// TIA Portal V20 export
// export: Created 2026-10-12T16:46:22.2661913Z, ExportSetting WithDefaults, DisplayName Totally Integrated Automation Portal, DisplayVersion V20 Update 6, DisplayName TIA Portal Openness, DisplayVersion V20 Update 6, DisplayName TIA Portal Version Control Interface, DisplayVersion V20 Update 6, DisplayName SINAMICS Startdrive Advanced, DisplayVersion V20 SP1 Update 2, DisplayName SINAMICS Startdrive G110M, G120, G120C, G120D, G120P, G115D, DisplayVersion V20 SP1 Update 2, DisplayName SINAMICS Startdrive G130, G150, S120, S150, SINAMICS MV, G220, S200, S210, DisplayVersion V20 SP1 Update 2, DisplayName STEP 7 Professional, DisplayVersion V20 Update 6, DisplayName STEP 7 Safety, DisplayVersion V20 Update 2, DisplayName WinCC Basic/Comfort/Advanced, DisplayVersion V20 Update 6, DisplayName WinCC Professional, DisplayVersion V20 Update 6, DisplayName WinCC Unified, DisplayVersion V20 Update 6
VAR_GLOBAL   // PLC tag table "KP8"
   "Maschinenleuchte orange ein P01" AT %Q1001.4 : Bool;
   "Maschinenleuchte gruen ein P01" AT %Q1001.5 : Bool;
   "Maschinenleuchte rot ein P01" AT %Q1001.6 : Bool;
   "Maschinenleuchte orange ein P02" AT %Q2001.4 : Bool;
   "Maschinenleuchte gruen ein P02" AT %Q2001.5 : Bool;
   "Maschinenleuchte rot ein P02" AT %Q2001.6 : Bool;
   "Maschinenleuchte orange ein P03" AT %Q3001.4 : Bool;
   "Maschinenleuchte gruen ein P03" AT %Q3001.5 : Bool;
   "Maschinenleuchte rot ein P03" AT %Q3001.6 : Bool;
   "Maschinenleuchte orange ein P04" AT %Q4001.4 : Bool;
   "Maschinenleuchte gruen ein P04" AT %Q4001.5 : Bool;
   "Maschinenleuchte rot ein P04" AT %Q4001.6 : Bool;
   "Maschinenleuchte orange ein P05" AT %Q5001.4 : Bool;
   "Maschinenleuchte gruen ein P05" AT %Q5001.5 : Bool;
   "Maschinenleuchte rot ein P05" AT %Q5001.6 : Bool;
   "Maschinenleuchte orange ein P06" AT %Q6001.4 : Bool;
   "Maschinenleuchte gruen ein P06" AT %Q6001.5 : Bool;
   "Maschinenleuchte rot ein P06" AT %Q6001.6 : Bool;
   "Maschinenleuchte orange ein P07" AT %Q7001.4 : Bool;
   "Maschinenleuchte gruen ein P07" AT %Q7001.5 : Bool;
   "Maschinenleuchte rot ein P07" AT %Q7001.6 : Bool;
   "Maschinenleuchte orange ein P08" AT %Q8001.4 : Bool;
   "Maschinenleuchte gruen ein P08" AT %Q8001.5 : Bool;
   "Maschinenleuchte rot ein P08" AT %Q8001.6 : Bool;
   "Maschinenleuchte orange ein P09" AT %Q9001.4 : Bool;
   "Maschinenleuchte gruen ein P09" AT %Q9001.5 : Bool;
   "Maschinenleuchte rot ein P09" AT %Q9001.6 : Bool;
   "Maschinenleuchte orange ein P10" AT %Q10001.4 : Bool;
   "Maschinenleuchte gruen ein P10" AT %Q10001.5 : Bool;
   "Maschinenleuchte rot ein P10" AT %Q10001.6 : Bool;
   "Maschinenleuchte orange ein P11" AT %Q11001.4 : Bool;
   "Maschinenleuchte gruen ein P11" AT %Q11001.5 : Bool;
   "Maschinenleuchte rot ein P11" AT %Q11001.6 : Bool;
   "Maschinenleuchte orange ein P12" AT %Q12001.4 : Bool;
   "Maschinenleuchte gruen ein P12" AT %Q12001.5 : Bool;
   "Maschinenleuchte rot ein P12" AT %Q12001.6 : Bool;
   "Maschinenleuchte orange ein P13" AT %Q13001.4 : Bool;
   "Maschinenleuchte gruen ein P13" AT %Q13001.5 : Bool;
   "Maschinenleuchte rot ein P13" AT %Q13001.6 : Bool;
   "Maschinenleuchte orange ein P14" AT %Q14001.4 : Bool;
   "Maschinenleuchte gruen ein P14" AT %Q14001.5 : Bool;
   "Maschinenleuchte rot ein P14" AT %Q14001.6 : Bool;
   "Maschinenleuchte orange ein P15" AT %Q15001.4 : Bool;
   "Maschinenleuchte gruen ein P15" AT %Q15001.5 : Bool;
   "Maschinenleuchte rot ein P15" AT %Q15001.6 : Bool;
   "Maschinenleuchte orange ein P16" AT %Q16001.4 : Bool;
   "Maschinenleuchte gruen ein P16" AT %Q16001.5 : Bool;
   "Maschinenleuchte rot ein P16" AT %Q16001.6 : Bool;
   "Maschinenleuchte orange ein P17" AT %Q17001.4 : Bool;
   "Maschinenleuchte gruen ein P17" AT %Q17001.5 : Bool;
   "Maschinenleuchte rot ein P17" AT %Q17001.6 : Bool;
   "Maschinenleuchte orange ein P18" AT %Q18001.4 : Bool;
   "Maschinenleuchte gruen ein P18" AT %Q18001.5 : Bool;
   "Maschinenleuchte rot ein P18" AT %Q18001.6 : Bool;
   "Maschinenleuchte orange ein P19" AT %Q19001.4 : Bool;
   "Maschinenleuchte gruen ein P19" AT %Q19001.5 : Bool;
   "Maschinenleuchte rot ein P19" AT %Q19001.6 : Bool;
   "Maschinenleuchte orange ein P20" AT %Q20001.4 : Bool;
   "Maschinenleuchte gruen ein P20" AT %Q20001.5 : Bool;
   "Maschinenleuchte rot ein P20" AT %Q20001.6 : Bool;
   "Maschinenleuchte orange ein P21" AT %Q21001.4 : Bool;
   "Maschinenleuchte gruen ein P21" AT %Q21001.5 : Bool;
   "Maschinenleuchte rot ein P21" AT %Q21001.6 : Bool;
   "Maschinenleuchte orange ein P22" AT %Q22001.4 : Bool;
   "Maschinenleuchte gruen ein P22" AT %Q22001.5 : Bool;
   "Maschinenleuchte rot ein P22" AT %Q22001.6 : Bool;
   "Maschinenleuchte orange ein P23" AT %Q23001.4 : Bool;
   "Maschinenleuchte gruen ein P23" AT %Q23001.5 : Bool;
   "Maschinenleuchte rot ein P23" AT %Q23001.6 : Bool;
   "Maschinenleuchte orange ein P24" AT %Q24001.4 : Bool;
   "Maschinenleuchte gruen ein P24" AT %Q24001.5 : Bool;
   "Maschinenleuchte rot ein P24" AT %Q24001.6 : Bool;
   "Maschinenleuchte orange ein P25" AT %Q25001.4 : Bool;
   "Maschinenleuchte gruen ein P25" AT %Q25001.5 : Bool;
   "Maschinenleuchte rot ein P25" AT %Q25001.6 : Bool;
   "Maschinenleuchte orange ein P26" AT %Q26001.4 : Bool;
   "Maschinenleuchte gruen ein P26" AT %Q26001.5 : Bool;
   "Maschinenleuchte rot ein P26" AT %Q26001.6 : Bool;
   "Maschinenleuchte orange ein P27" AT %Q27001.4 : Bool;
   "Maschinenleuchte gruen ein P27" AT %Q27001.5 : Bool;
   "Maschinenleuchte rot ein P27" AT %Q27001.6 : Bool;
   "Maschinenleuchte orange ein P28" AT %Q28001.4 : Bool;
   "Maschinenleuchte gruen ein P28" AT %Q28001.5 : Bool;
   "Maschinenleuchte rot ein P28" AT %Q28001.6 : Bool;
END_VAR
